PROGRAM main
  VAR
    Button AT %QX0.0 : BOOL;
    MOTOR AT %QX0.1 : BOOL;
    PULSE AT %QX0.2 : BOOL;
    RESET_ALL AT %QX0.3 : BOOL;
    WEIGHT_SEN AT %MW0 : INT;
    COUNT AT %MW1 : INT;
    BIG_BOX_COUNT AT %MW2 : INT;
    MEDIUM_BOX_COUNT AT %MW3 : INT;
    SMAll_BOX_COUNT AT %MW4 : INT;
    isbig AT %MX0.0 : BOOL;
    is_medium AT %MX0.1 : BOOL;
    is_small AT %MX0.2 : BOOL;
    CTU0 : CTU;
    less_than_10 : BOOL;
    greather_than_5 : BOOL;
    CTU1 : CTU;
    CTU2 : CTU;
    CTU3 : CTU;
    CTU4 : CTU;
    TON0 : TON;
    AllocateA : BOOL;
    TON1 : TON;
    TON2 : TON;
    AllocateB : BOOL;
    AllocateC : BOOL;
  END_VAR

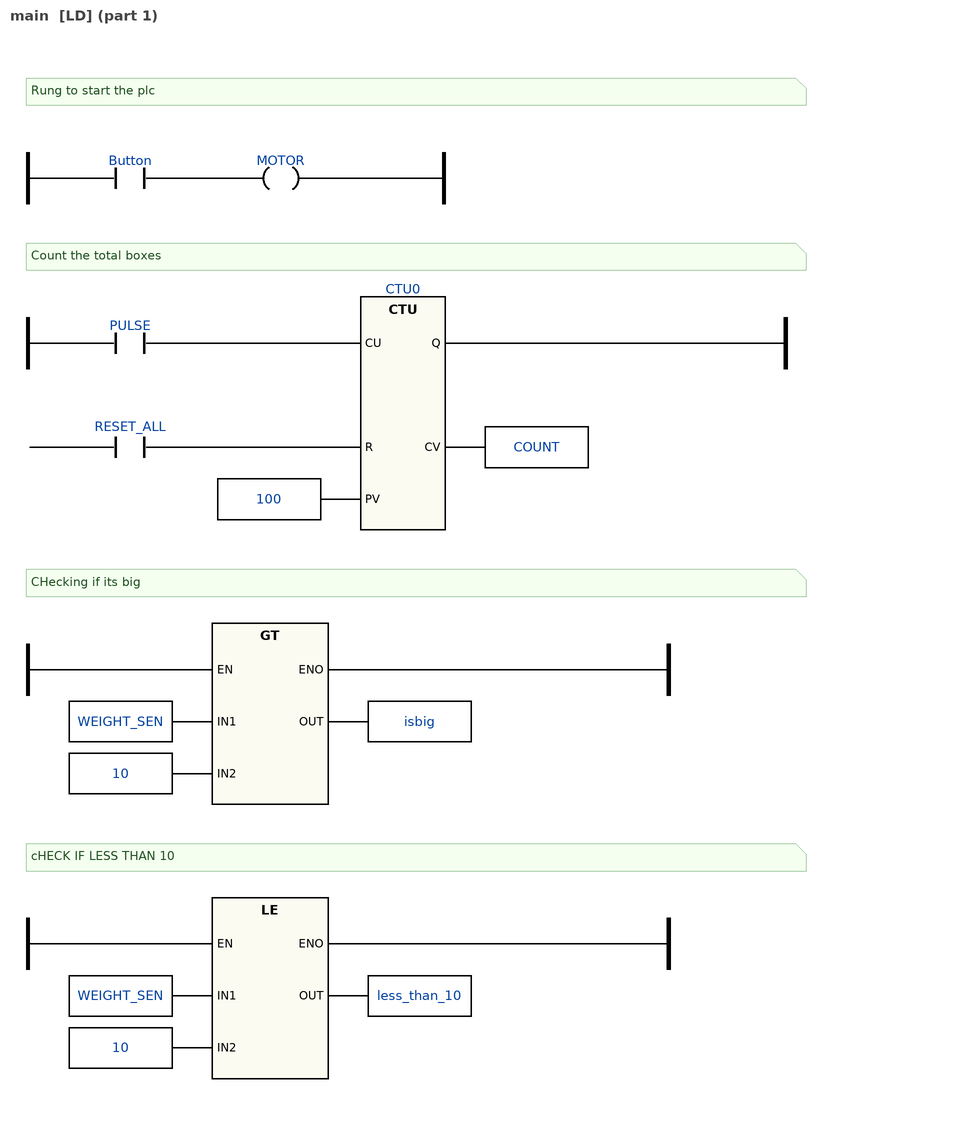
(* LD diagram, written out as Structured Text *)
(* Rung to start the plc *)
MOTOR := Button;
(* Count the total boxes *)
CTU0(CU := PULSE, R := RESET_ALL, PV := 100);
COUNT := CTU0.CV;
(* CHecking if its big *)
isbig := WEIGHT_SEN > 10;
(* cHECK IF LESS THAN 10 *)
less_than_10 := WEIGHT_SEN <= 10;
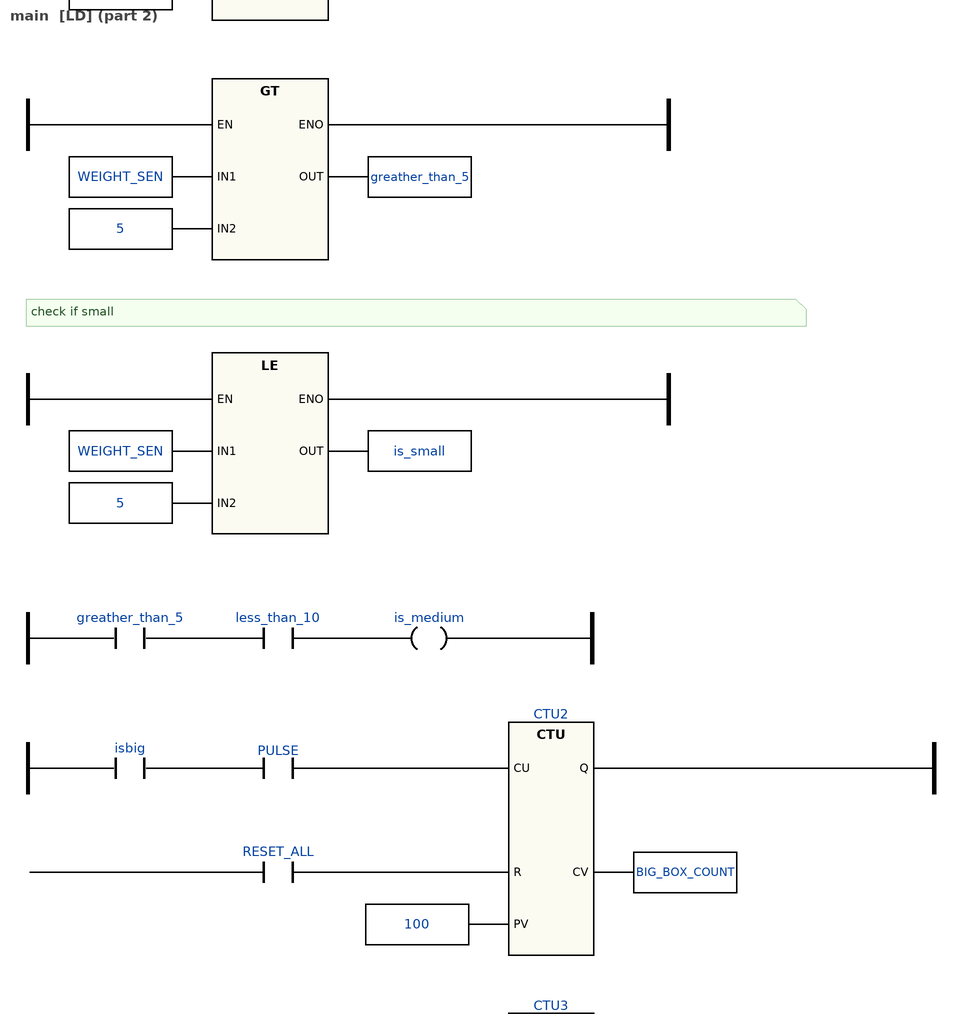
greather_than_5 := WEIGHT_SEN > 5;
(* check if small *)
is_small := WEIGHT_SEN <= 5;
is_medium := greather_than_5 AND less_than_10;
CTU2(CU := isbig AND PULSE, R := RESET_ALL, PV := 100);
BIG_BOX_COUNT := CTU2.CV;
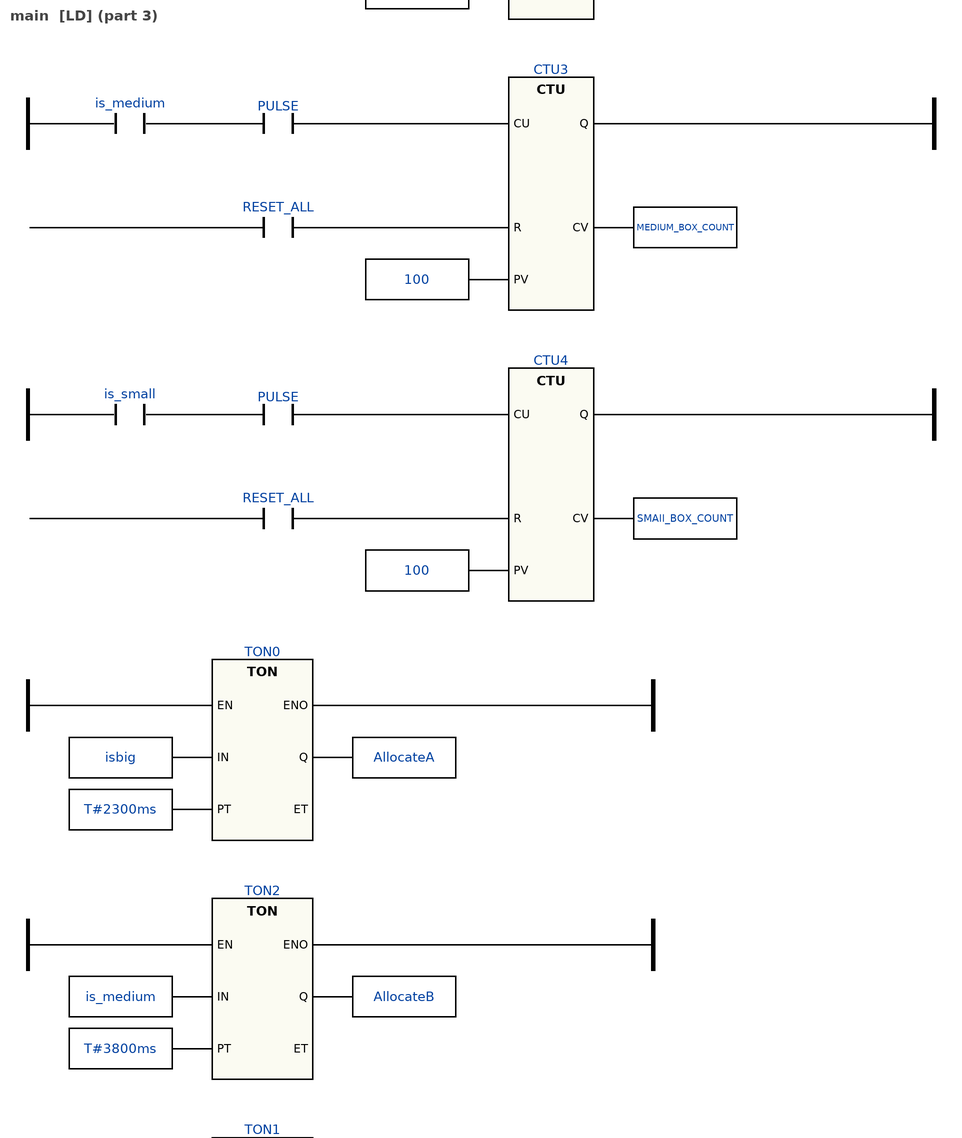
CTU3(CU := is_medium AND PULSE, R := RESET_ALL, PV := 100);
MEDIUM_BOX_COUNT := CTU3.CV;
CTU4(CU := is_small AND PULSE, R := RESET_ALL, PV := 100);
SMAll_BOX_COUNT := CTU4.CV;
TON0(IN := isbig, PT := T#2300ms);
AllocateA := TON0.Q;
TON2(IN := is_medium, PT := T#3800ms);
AllocateB := TON2.Q;
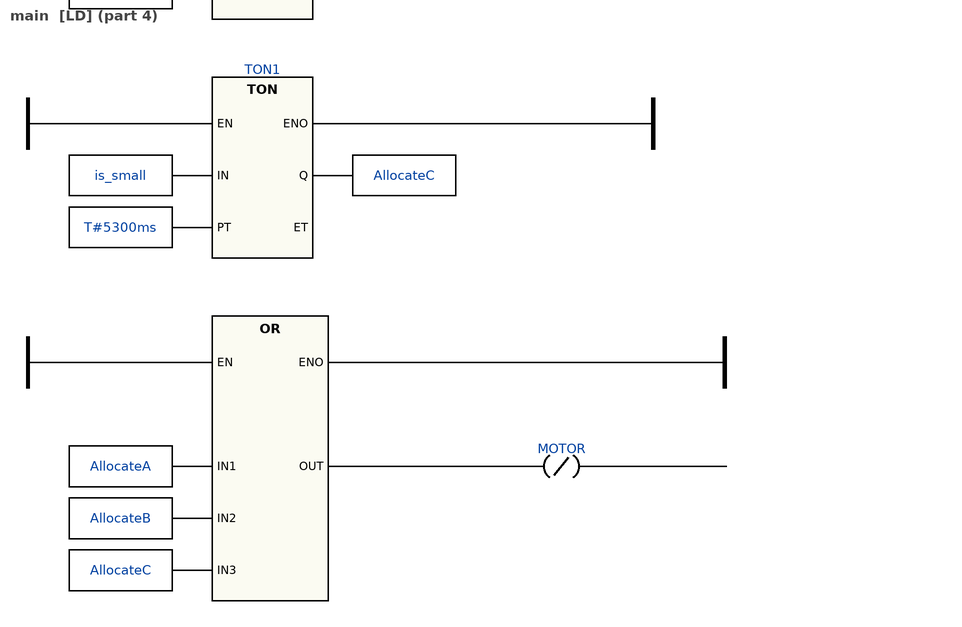
TON1(IN := is_small, PT := T#5300ms);
AllocateC := TON1.Q;
MOTOR := NOT (AllocateA OR AllocateB OR AllocateC);
END_PROGRAM
